(* Schneider Machine Expert - Basic project Case07, file version 2.9.0.0 *)
(* ProjectInformations: Name=New project *)

HARDWARE
  Cpu 0: TM221M16R/G
  EthernetConfiguration: NetworkName=M221, IpAllocationMode=FixedAddress, IpAddress=0.0.0.0, SubnetMask=0.0.0.0
  SerialLineConfiguration: Baud=Baud19200, Parity=ParityEven, DataBits=DataBits8, StopBits=StopBits1, PhysicalMedium=PhysicalMediumRs485, TransmissionMode=TransmissionModeModbusRtu, SlaveId=1, Addressing=SlaveAddressing
  MastTask: UsePeriodScanMode=false, PeriodScan=100
  FastTask: Period=255
  CpuBehavior: StartingMode=StartAsPreviousState, AutoSaveRamOnEeprom=true, WatchdogPeriod=250

SYMBOLS  (address, symbol, comment, settings)
  %M10      Initialised
  %M11      Stage0
  %M12      Stage1
  %M13      Stage2
  %M14      Stage3
  %M15      Stage4
  %M16      Stage5
  %M17      Stage6
  %M18      Stage7
  %M19      Hold0
  %M20      Hold1
  %M21      Hold2
  %M22      Hold3
  %M23      Hold4
  %M24      Hold5
  %M25      Hold6
  %M26      Hold7
  %M27      Advance0
  %M28      Advance1
  %M29      Advance2
  %M30      Advance3
  %M31      Advance4
  %M32      Advance5
  %M33      Advance6
  %M34      Advance7
  %M35      NSGreenPermit
  %M36      NSYellowPermit
  %M37      EWGreenPermit
  %M38      EWYellowPermit
  %M39      PedGreenPermit
  %M100     NorthRed
  %M101     NorthYellow
  %M102     NorthGreen
  %M103     SouthRed
  %M104     SouthYellow
  %M105     SouthGreen
  %M106     EastRed
  %M107     EastYellow
  %M108     EastGreen
  %M109     WestRed
  %M110     WestYellow
  %M111     WestGreen
  %M112     PedRed
  %M113     PedGreen
  %TM0        [Preset=2, Base=OneSecond]
  %TM1        [Preset=10, Base=OneSecond]
  %TM2        [Preset=3, Base=OneSecond]
  %TM3        [Preset=2, Base=OneSecond]
  %TM4        [Preset=10, Base=OneSecond]
  %TM5        [Preset=3, Base=OneSecond]
  %TM6        [Preset=2, Base=OneSecond]
  %TM7        [Preset=5, Base=OneSecond]

POU New POU
  (* SectionNumber=1 *)

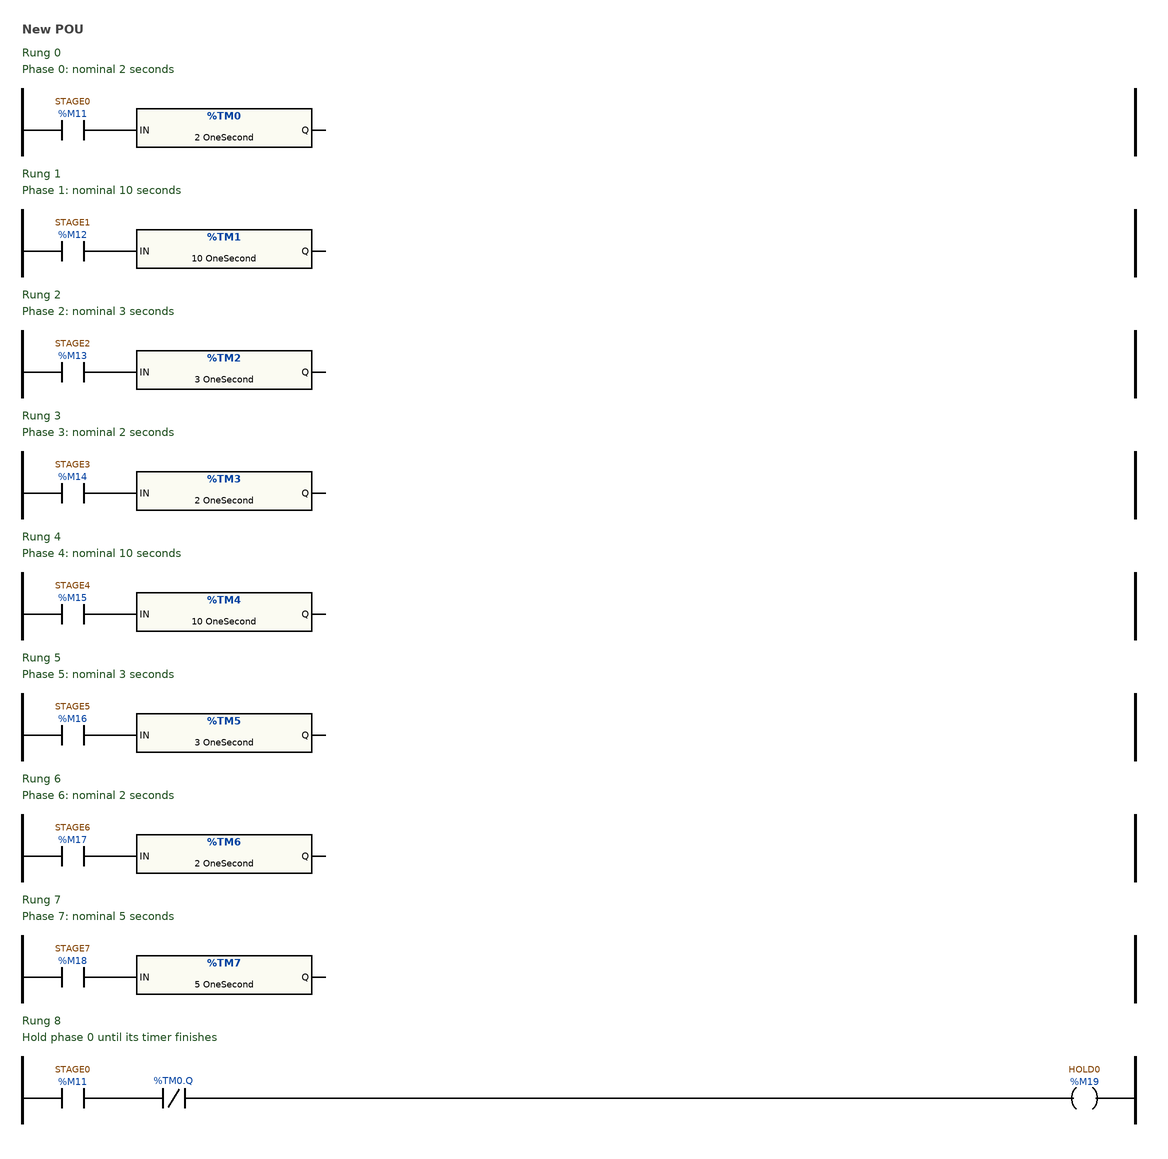

// Rung 0
// Phase 0: nominal 2 seconds
  BLK %TM0
  LD %M11                 (* Stage0 *)
  IN
  END_BLK
  // as ST:
  //   %TM0(IN := Stage0);

// Rung 1
// Phase 1: nominal 10 seconds
  BLK %TM1
  LD %M12                 (* Stage1 *)
  IN
  END_BLK
  // as ST:
  //   %TM1(IN := Stage1);

// Rung 2
// Phase 2: nominal 3 seconds
  BLK %TM2
  LD %M13                 (* Stage2 *)
  IN
  END_BLK
  // as ST:
  //   %TM2(IN := Stage2);

// Rung 3
// Phase 3: nominal 2 seconds
  BLK %TM3
  LD %M14                 (* Stage3 *)
  IN
  END_BLK
  // as ST:
  //   %TM3(IN := Stage3);

// Rung 4
// Phase 4: nominal 10 seconds
  BLK %TM4
  LD %M15                 (* Stage4 *)
  IN
  END_BLK
  // as ST:
  //   %TM4(IN := Stage4);

// Rung 5
// Phase 5: nominal 3 seconds
  BLK %TM5
  LD %M16                 (* Stage5 *)
  IN
  END_BLK
  // as ST:
  //   %TM5(IN := Stage5);

// Rung 6
// Phase 6: nominal 2 seconds
  BLK %TM6
  LD %M17                 (* Stage6 *)
  IN
  END_BLK
  // as ST:
  //   %TM6(IN := Stage6);

// Rung 7
// Phase 7: nominal 5 seconds
  BLK %TM7
  LD %M18                 (* Stage7 *)
  IN
  END_BLK
  // as ST:
  //   %TM7(IN := Stage7);

// Rung 8
// Hold phase 0 until its timer finishes
  LD %M11                 (* Stage0 *)
  ANDN %TM0.Q
  ST %M19                 (* Hold0 *)
  // as ST:
  //   Hold0 := Stage0 AND NOT %TM0.Q;

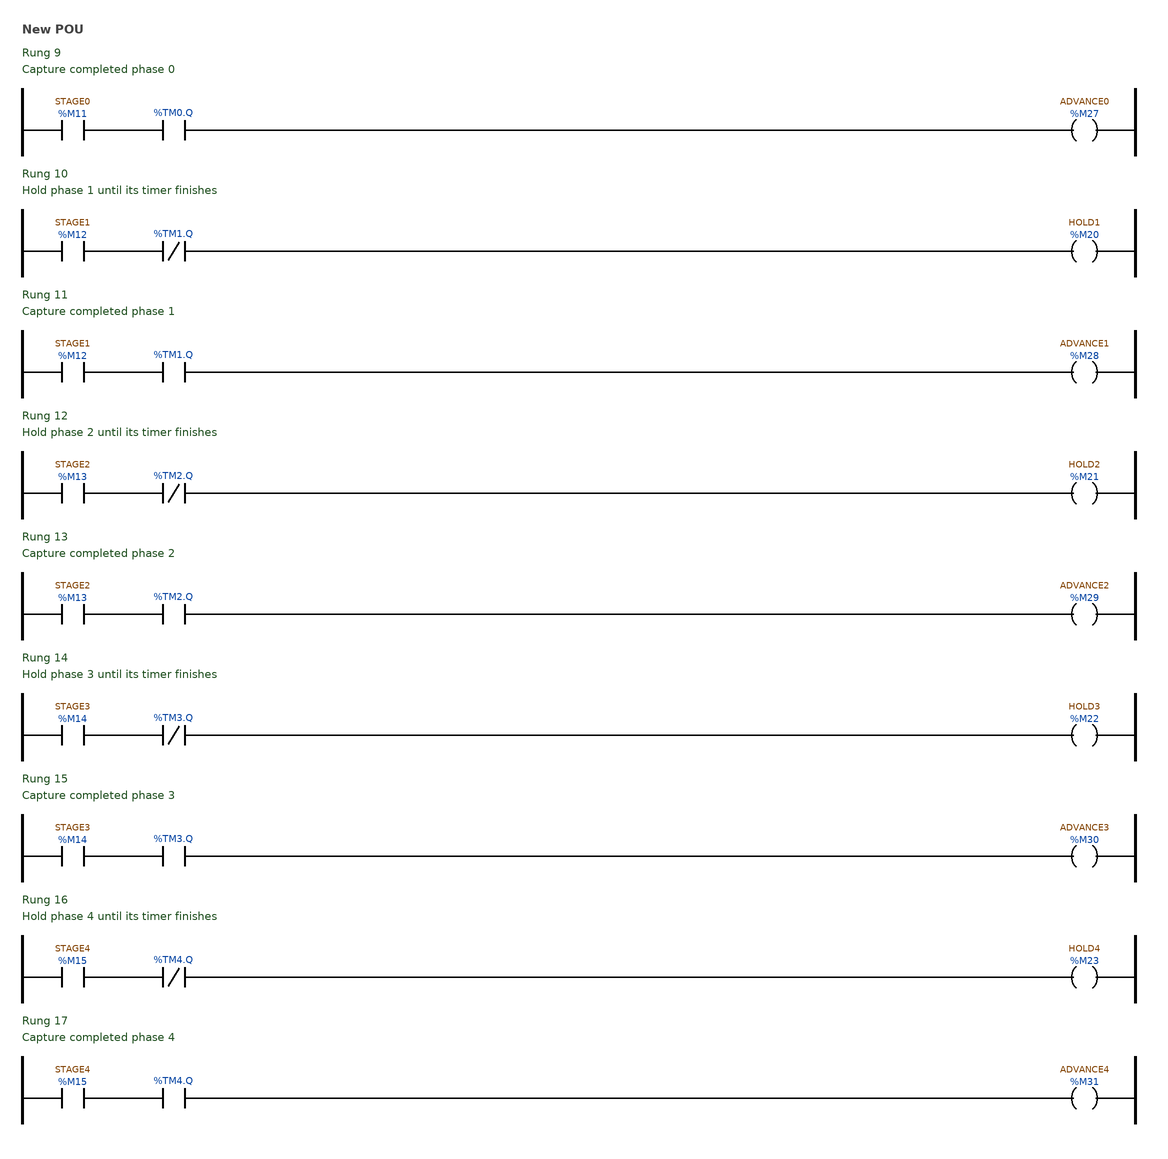

// Rung 9
// Capture completed phase 0
  LD %M11                 (* Stage0 *)
  AND %TM0.Q
  ST %M27                 (* Advance0 *)
  // as ST:
  //   Advance0 := Stage0 AND %TM0.Q;

// Rung 10
// Hold phase 1 until its timer finishes
  LD %M12                 (* Stage1 *)
  ANDN %TM1.Q
  ST %M20                 (* Hold1 *)
  // as ST:
  //   Hold1 := Stage1 AND NOT %TM1.Q;

// Rung 11
// Capture completed phase 1
  LD %M12                 (* Stage1 *)
  AND %TM1.Q
  ST %M28                 (* Advance1 *)
  // as ST:
  //   Advance1 := Stage1 AND %TM1.Q;

// Rung 12
// Hold phase 2 until its timer finishes
  LD %M13                 (* Stage2 *)
  ANDN %TM2.Q
  ST %M21                 (* Hold2 *)
  // as ST:
  //   Hold2 := Stage2 AND NOT %TM2.Q;

// Rung 13
// Capture completed phase 2
  LD %M13                 (* Stage2 *)
  AND %TM2.Q
  ST %M29                 (* Advance2 *)
  // as ST:
  //   Advance2 := Stage2 AND %TM2.Q;

// Rung 14
// Hold phase 3 until its timer finishes
  LD %M14                 (* Stage3 *)
  ANDN %TM3.Q
  ST %M22                 (* Hold3 *)
  // as ST:
  //   Hold3 := Stage3 AND NOT %TM3.Q;

// Rung 15
// Capture completed phase 3
  LD %M14                 (* Stage3 *)
  AND %TM3.Q
  ST %M30                 (* Advance3 *)
  // as ST:
  //   Advance3 := Stage3 AND %TM3.Q;

// Rung 16
// Hold phase 4 until its timer finishes
  LD %M15                 (* Stage4 *)
  ANDN %TM4.Q
  ST %M23                 (* Hold4 *)
  // as ST:
  //   Hold4 := Stage4 AND NOT %TM4.Q;

// Rung 17
// Capture completed phase 4
  LD %M15                 (* Stage4 *)
  AND %TM4.Q
  ST %M31                 (* Advance4 *)
  // as ST:
  //   Advance4 := Stage4 AND %TM4.Q;

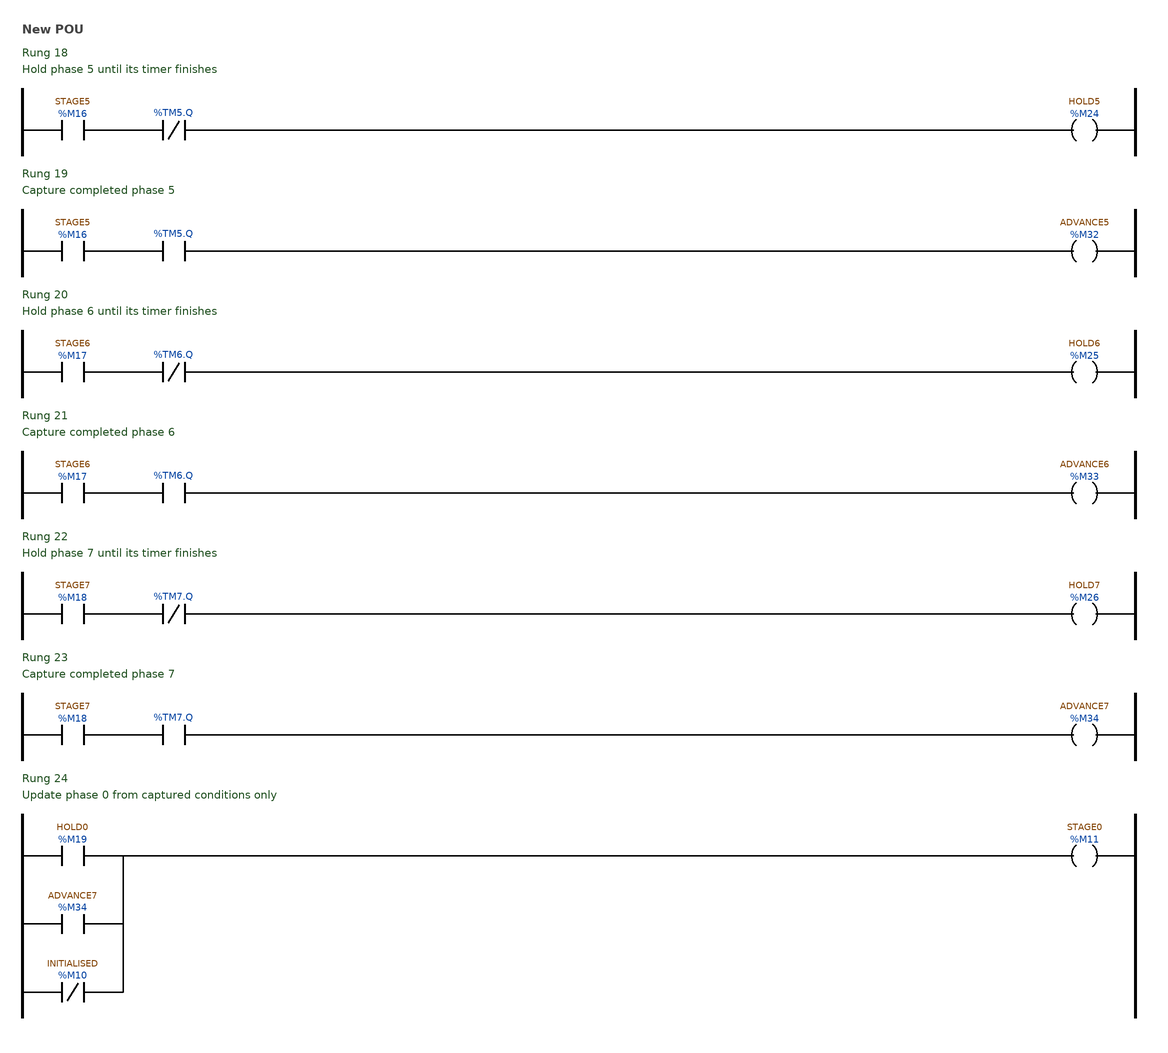

// Rung 18
// Hold phase 5 until its timer finishes
  LD %M16                 (* Stage5 *)
  ANDN %TM5.Q
  ST %M24                 (* Hold5 *)
  // as ST:
  //   Hold5 := Stage5 AND NOT %TM5.Q;

// Rung 19
// Capture completed phase 5
  LD %M16                 (* Stage5 *)
  AND %TM5.Q
  ST %M32                 (* Advance5 *)
  // as ST:
  //   Advance5 := Stage5 AND %TM5.Q;

// Rung 20
// Hold phase 6 until its timer finishes
  LD %M17                 (* Stage6 *)
  ANDN %TM6.Q
  ST %M25                 (* Hold6 *)
  // as ST:
  //   Hold6 := Stage6 AND NOT %TM6.Q;

// Rung 21
// Capture completed phase 6
  LD %M17                 (* Stage6 *)
  AND %TM6.Q
  ST %M33                 (* Advance6 *)
  // as ST:
  //   Advance6 := Stage6 AND %TM6.Q;

// Rung 22
// Hold phase 7 until its timer finishes
  LD %M18                 (* Stage7 *)
  ANDN %TM7.Q
  ST %M26                 (* Hold7 *)
  // as ST:
  //   Hold7 := Stage7 AND NOT %TM7.Q;

// Rung 23
// Capture completed phase 7
  LD %M18                 (* Stage7 *)
  AND %TM7.Q
  ST %M34                 (* Advance7 *)
  // as ST:
  //   Advance7 := Stage7 AND %TM7.Q;

// Rung 24
// Update phase 0 from captured conditions only
  LD %M19                 (* Hold0 *)
  OR %M34                 (* Advance7 *)
  ORN %M10                (* Initialised *)
  ST %M11                 (* Stage0 *)
  // as ST:
  //   Stage0 := Hold0 OR Advance7 OR NOT Initialised;

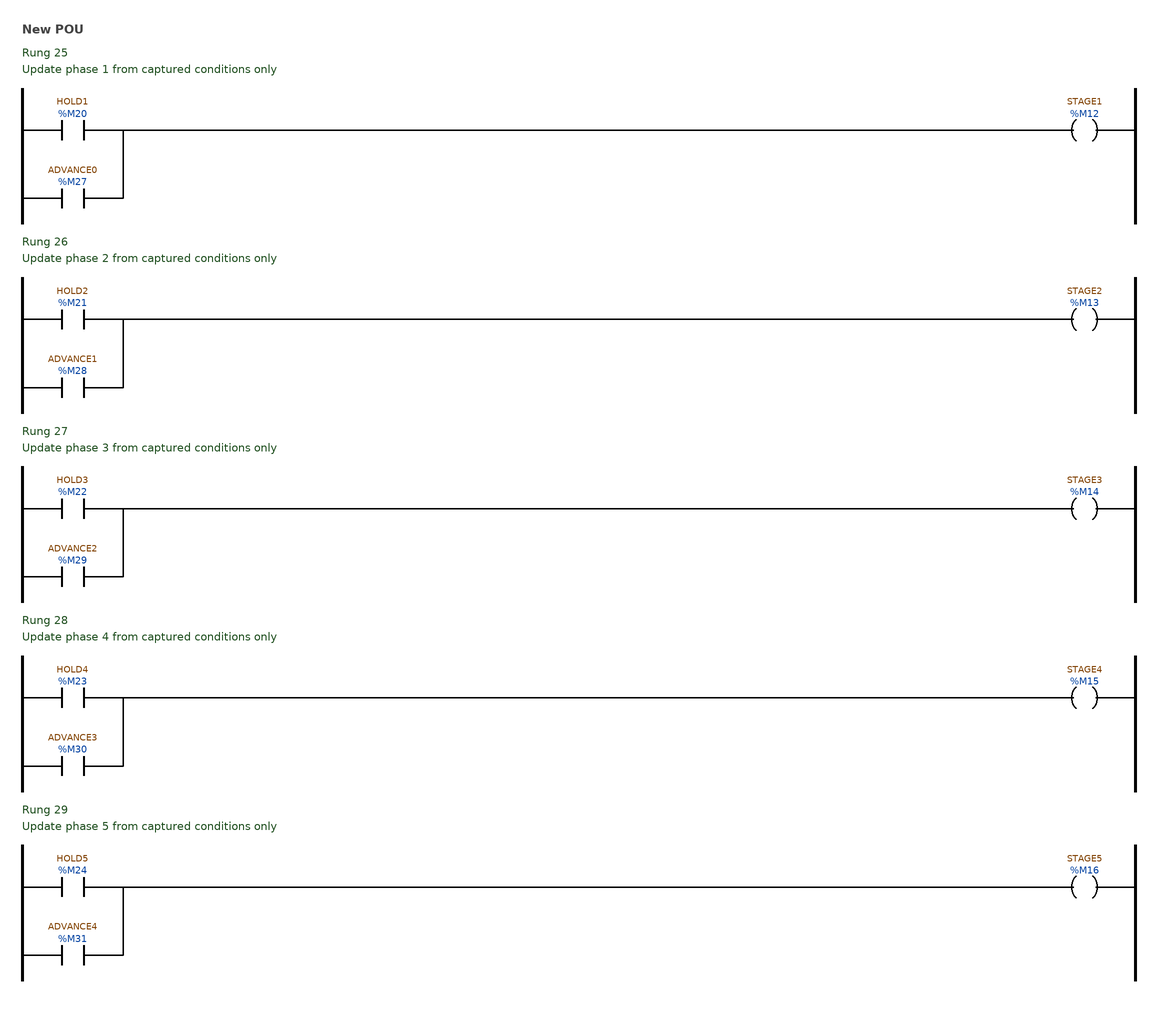

// Rung 25
// Update phase 1 from captured conditions only
  LD %M20                 (* Hold1 *)
  OR %M27                 (* Advance0 *)
  ST %M12                 (* Stage1 *)
  // as ST:
  //   Stage1 := Hold1 OR Advance0;

// Rung 26
// Update phase 2 from captured conditions only
  LD %M21                 (* Hold2 *)
  OR %M28                 (* Advance1 *)
  ST %M13                 (* Stage2 *)
  // as ST:
  //   Stage2 := Hold2 OR Advance1;

// Rung 27
// Update phase 3 from captured conditions only
  LD %M22                 (* Hold3 *)
  OR %M29                 (* Advance2 *)
  ST %M14                 (* Stage3 *)
  // as ST:
  //   Stage3 := Hold3 OR Advance2;

// Rung 28
// Update phase 4 from captured conditions only
  LD %M23                 (* Hold4 *)
  OR %M30                 (* Advance3 *)
  ST %M15                 (* Stage4 *)
  // as ST:
  //   Stage4 := Hold4 OR Advance3;

// Rung 29
// Update phase 5 from captured conditions only
  LD %M24                 (* Hold5 *)
  OR %M31                 (* Advance4 *)
  ST %M16                 (* Stage5 *)
  // as ST:
  //   Stage5 := Hold5 OR Advance4;

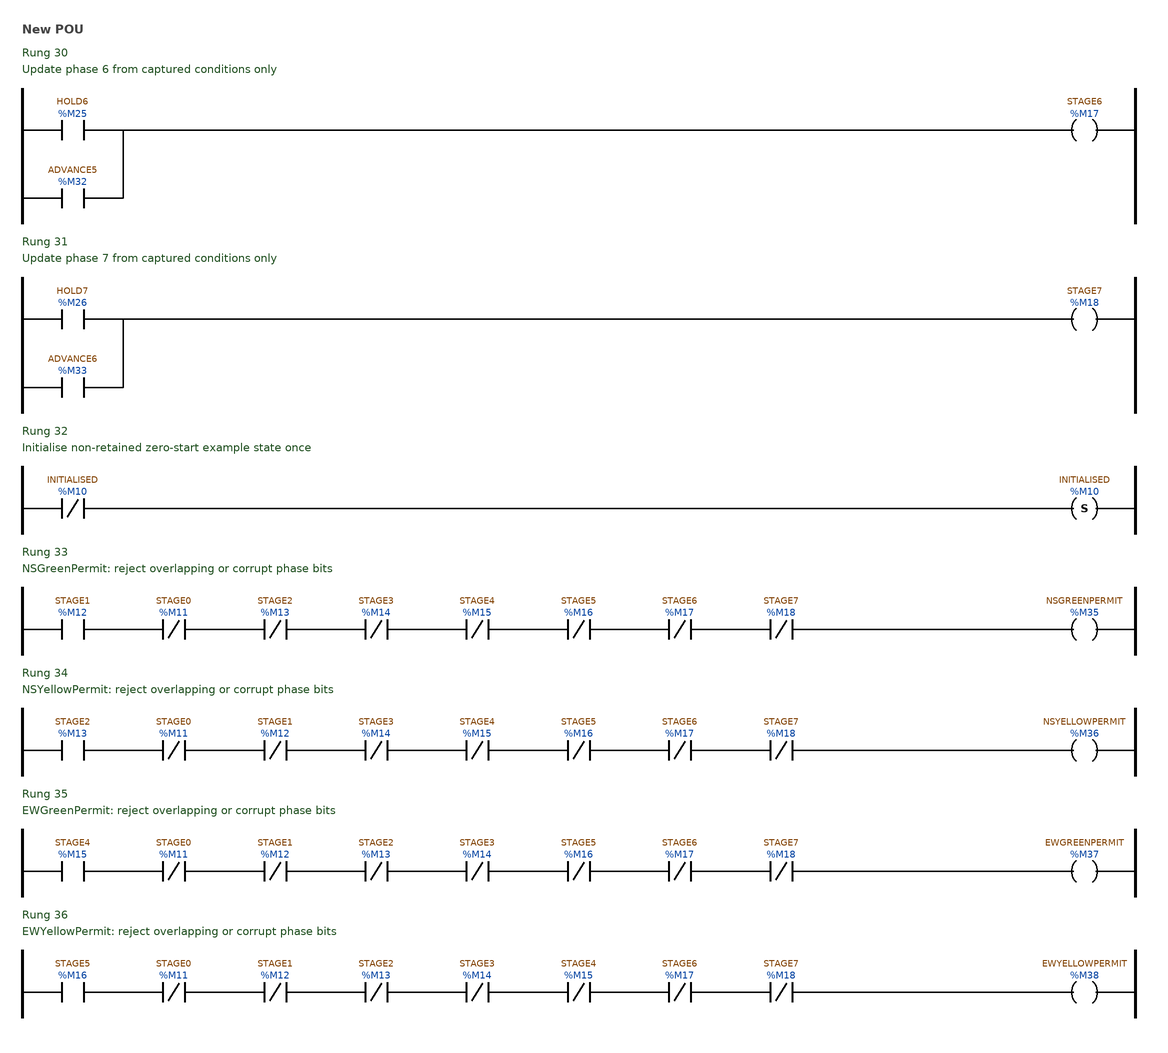

// Rung 30
// Update phase 6 from captured conditions only
  LD %M25                 (* Hold6 *)
  OR %M32                 (* Advance5 *)
  ST %M17                 (* Stage6 *)
  // as ST:
  //   Stage6 := Hold6 OR Advance5;

// Rung 31
// Update phase 7 from captured conditions only
  LD %M26                 (* Hold7 *)
  OR %M33                 (* Advance6 *)
  ST %M18                 (* Stage7 *)
  // as ST:
  //   Stage7 := Hold7 OR Advance6;

// Rung 32
// Initialise non-retained zero-start example state once
  LDN %M10                (* Initialised *)
  S %M10                  (* Initialised *)
  // as ST:
  //   IF NOT Initialised THEN Initialised := TRUE; END_IF;

// Rung 33
// NSGreenPermit: reject overlapping or corrupt phase bits
  LD %M12                 (* Stage1 *)
  ANDN %M11               (* Stage0 *)
  ANDN %M13               (* Stage2 *)
  ANDN %M14               (* Stage3 *)
  ANDN %M15               (* Stage4 *)
  ANDN %M16               (* Stage5 *)
  ANDN %M17               (* Stage6 *)
  ANDN %M18               (* Stage7 *)
  ST %M35                 (* NSGreenPermit *)
  // as ST:
  //   NSGreenPermit := Stage1 AND NOT Stage0 AND NOT Stage2 AND NOT Stage3 AND NOT Stage4 AND NOT Stage5 AND NOT Stage6 AND NOT Stage7;

// Rung 34
// NSYellowPermit: reject overlapping or corrupt phase bits
  LD %M13                 (* Stage2 *)
  ANDN %M11               (* Stage0 *)
  ANDN %M12               (* Stage1 *)
  ANDN %M14               (* Stage3 *)
  ANDN %M15               (* Stage4 *)
  ANDN %M16               (* Stage5 *)
  ANDN %M17               (* Stage6 *)
  ANDN %M18               (* Stage7 *)
  ST %M36                 (* NSYellowPermit *)
  // as ST:
  //   NSYellowPermit := Stage2 AND NOT Stage0 AND NOT Stage1 AND NOT Stage3 AND NOT Stage4 AND NOT Stage5 AND NOT Stage6 AND NOT Stage7;

// Rung 35
// EWGreenPermit: reject overlapping or corrupt phase bits
  LD %M15                 (* Stage4 *)
  ANDN %M11               (* Stage0 *)
  ANDN %M12               (* Stage1 *)
  ANDN %M13               (* Stage2 *)
  ANDN %M14               (* Stage3 *)
  ANDN %M16               (* Stage5 *)
  ANDN %M17               (* Stage6 *)
  ANDN %M18               (* Stage7 *)
  ST %M37                 (* EWGreenPermit *)
  // as ST:
  //   EWGreenPermit := Stage4 AND NOT Stage0 AND NOT Stage1 AND NOT Stage2 AND NOT Stage3 AND NOT Stage5 AND NOT Stage6 AND NOT Stage7;

// Rung 36
// EWYellowPermit: reject overlapping or corrupt phase bits
  LD %M16                 (* Stage5 *)
  ANDN %M11               (* Stage0 *)
  ANDN %M12               (* Stage1 *)
  ANDN %M13               (* Stage2 *)
  ANDN %M14               (* Stage3 *)
  ANDN %M15               (* Stage4 *)
  ANDN %M17               (* Stage6 *)
  ANDN %M18               (* Stage7 *)
  ST %M38                 (* EWYellowPermit *)
  // as ST:
  //   EWYellowPermit := Stage5 AND NOT Stage0 AND NOT Stage1 AND NOT Stage2 AND NOT Stage3 AND NOT Stage4 AND NOT Stage6 AND NOT Stage7;

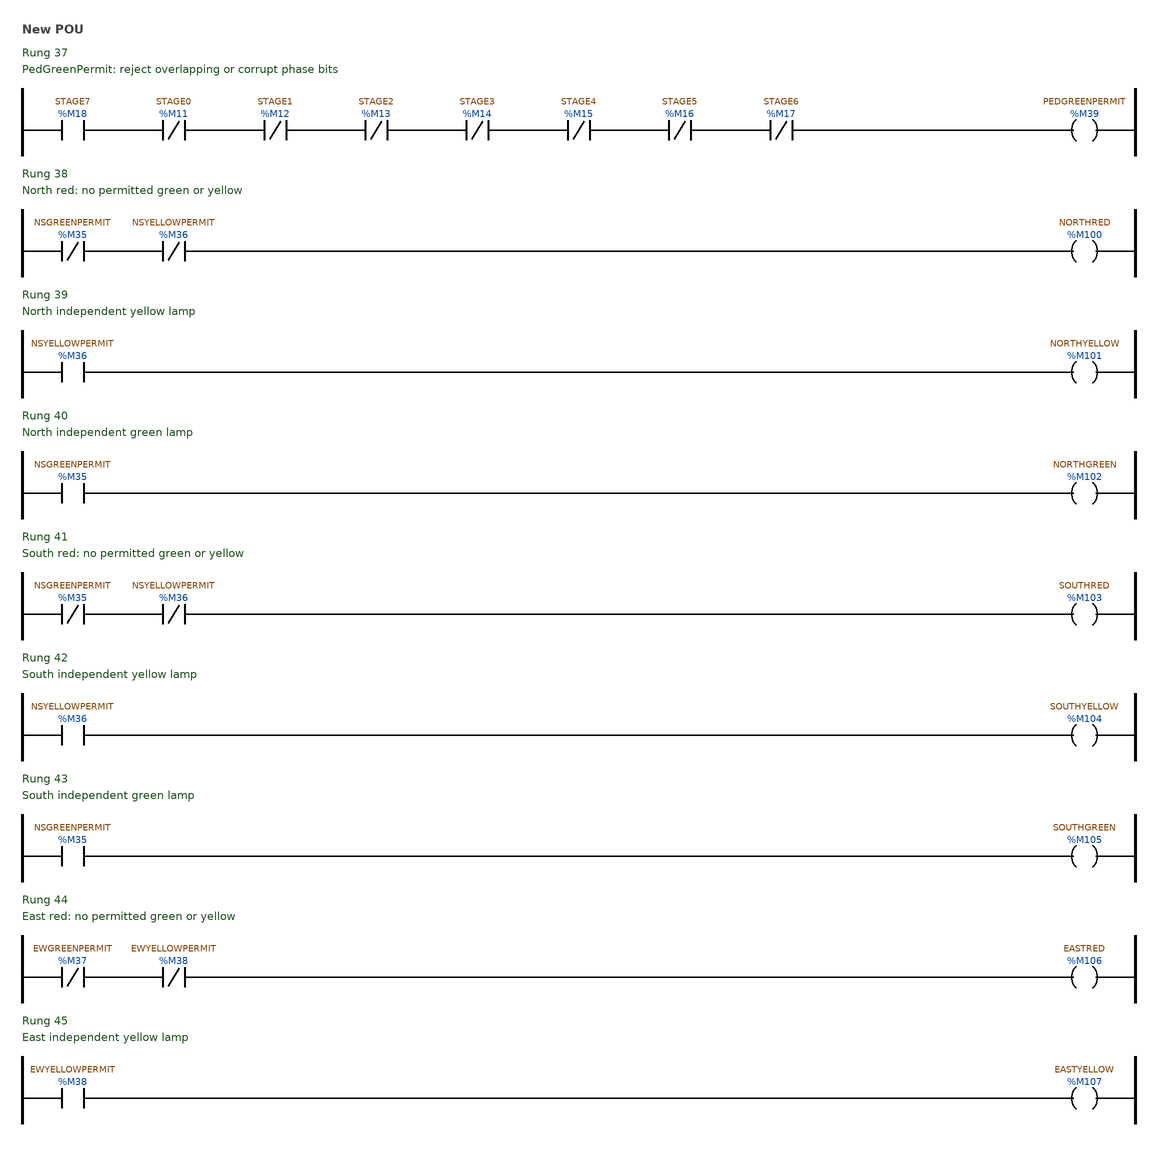

// Rung 37
// PedGreenPermit: reject overlapping or corrupt phase bits
  LD %M18                 (* Stage7 *)
  ANDN %M11               (* Stage0 *)
  ANDN %M12               (* Stage1 *)
  ANDN %M13               (* Stage2 *)
  ANDN %M14               (* Stage3 *)
  ANDN %M15               (* Stage4 *)
  ANDN %M16               (* Stage5 *)
  ANDN %M17               (* Stage6 *)
  ST %M39                 (* PedGreenPermit *)
  // as ST:
  //   PedGreenPermit := Stage7 AND NOT Stage0 AND NOT Stage1 AND NOT Stage2 AND NOT Stage3 AND NOT Stage4 AND NOT Stage5 AND NOT Stage6;

// Rung 38
// North red: no permitted green or yellow
  LDN %M35                (* NSGreenPermit *)
  ANDN %M36               (* NSYellowPermit *)
  ST %M100                (* NorthRed *)
  // as ST:
  //   NorthRed := NOT NSGreenPermit AND NOT NSYellowPermit;

// Rung 39
// North independent yellow lamp
  LD %M36                 (* NSYellowPermit *)
  ST %M101                (* NorthYellow *)
  // as ST:
  //   NorthYellow := NSYellowPermit;

// Rung 40
// North independent green lamp
  LD %M35                 (* NSGreenPermit *)
  ST %M102                (* NorthGreen *)
  // as ST:
  //   NorthGreen := NSGreenPermit;

// Rung 41
// South red: no permitted green or yellow
  LDN %M35                (* NSGreenPermit *)
  ANDN %M36               (* NSYellowPermit *)
  ST %M103                (* SouthRed *)
  // as ST:
  //   SouthRed := NOT NSGreenPermit AND NOT NSYellowPermit;

// Rung 42
// South independent yellow lamp
  LD %M36                 (* NSYellowPermit *)
  ST %M104                (* SouthYellow *)
  // as ST:
  //   SouthYellow := NSYellowPermit;

// Rung 43
// South independent green lamp
  LD %M35                 (* NSGreenPermit *)
  ST %M105                (* SouthGreen *)
  // as ST:
  //   SouthGreen := NSGreenPermit;

// Rung 44
// East red: no permitted green or yellow
  LDN %M37                (* EWGreenPermit *)
  ANDN %M38               (* EWYellowPermit *)
  ST %M106                (* EastRed *)
  // as ST:
  //   EastRed := NOT EWGreenPermit AND NOT EWYellowPermit;

// Rung 45
// East independent yellow lamp
  LD %M38                 (* EWYellowPermit *)
  ST %M107                (* EastYellow *)
  // as ST:
  //   EastYellow := EWYellowPermit;

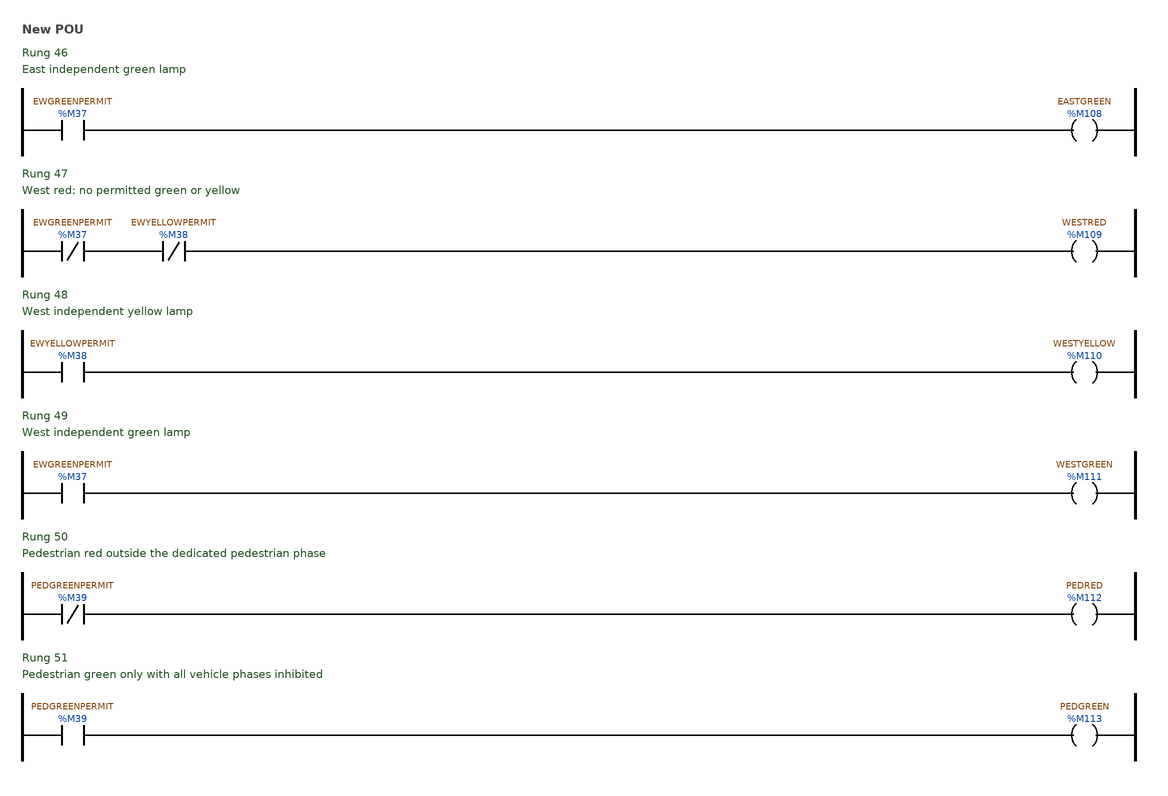

// Rung 46
// East independent green lamp
  LD %M37                 (* EWGreenPermit *)
  ST %M108                (* EastGreen *)
  // as ST:
  //   EastGreen := EWGreenPermit;

// Rung 47
// West red: no permitted green or yellow
  LDN %M37                (* EWGreenPermit *)
  ANDN %M38               (* EWYellowPermit *)
  ST %M109                (* WestRed *)
  // as ST:
  //   WestRed := NOT EWGreenPermit AND NOT EWYellowPermit;

// Rung 48
// West independent yellow lamp
  LD %M38                 (* EWYellowPermit *)
  ST %M110                (* WestYellow *)
  // as ST:
  //   WestYellow := EWYellowPermit;

// Rung 49
// West independent green lamp
  LD %M37                 (* EWGreenPermit *)
  ST %M111                (* WestGreen *)
  // as ST:
  //   WestGreen := EWGreenPermit;

// Rung 50
// Pedestrian red outside the dedicated pedestrian phase
  LDN %M39                (* PedGreenPermit *)
  ST %M112                (* PedRed *)
  // as ST:
  //   PedRed := NOT PedGreenPermit;

// Rung 51
// Pedestrian green only with all vehicle phases inhibited
  LD %M39                 (* PedGreenPermit *)
  ST %M113                (* PedGreen *)
  // as ST:
  //   PedGreen := PedGreenPermit;
